TYPE "ST_PressDemoStationCfg"
VERSION : 0.1
   STRUCT
      SchemaVersion : UInt := 1;
      RequireTwoHandStart : Bool := TRUE;
      TransferSettleTime : Time := T#200MS;
      PressSettleTime : Time := T#300MS;
   END_STRUCT;

END_TYPE

